FUNCTION_BLOCK FB_PackagingCounter (* Migrated from IEC 61131-3 ST *)
  (* Standard: 61499-2 *)
  (* Version 1.0, 2026-11-06, st2fb *)
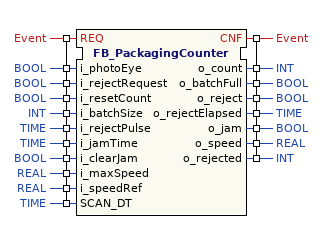
  EVENT_INPUT
    REQ WITH i_photoEye, i_rejectRequest, i_resetCount, i_batchSize, i_rejectPulse, i_jamTime, i_clearJam, i_maxSpeed, i_speedRef, SCAN_DT;
  END_EVENT
  EVENT_OUTPUT
    CNF WITH o_count, o_batchFull, o_reject, o_rejectElapsed, o_jam, o_speed, o_rejected;
  END_EVENT
  VAR_INPUT
    i_photoEye : BOOL;
    i_rejectRequest : BOOL;
    i_resetCount : BOOL;
    i_batchSize : INT;
    i_rejectPulse : TIME;
    i_jamTime : TIME;
    i_clearJam : BOOL;
    i_maxSpeed : REAL;
    i_speedRef : REAL;
    SCAN_DT : TIME;
  END_VAR
  VAR_OUTPUT
    o_count : INT;
    o_batchFull : BOOL;
    o_reject : BOOL;
    o_rejectElapsed : TIME;
    o_jam : BOOL;
    o_speed : REAL;
    o_rejected : INT;
  END_VAR
  VAR
    statEyePrev : BOOL := FALSE;
    statRequestPrev : BOOL := FALSE;
    statRejectPrev : BOOL := FALSE;
    statRejectPreset : TIME := T#0s;
    statJamPreset : TIME := T#0s;
    tempCartonEdge : BOOL := FALSE;
    tempRejectEdge : BOOL := FALSE;
    ST2FB_NOW : TIME := T#0s;
    RP_IN : BOOL := FALSE;
    RP_PT : TIME := T#0s;
    RP_Q : BOOL := FALSE;
    RP_ET : TIME := T#0s;
    RP_STATE : INT := 0;
    RP_PREV_IN : BOOL := FALSE;
    RP_START_TIME : TIME := T#0s;
    JT_IN : BOOL := FALSE;
    JT_PT : TIME := T#0s;
    JT_Q : BOOL := FALSE;
    JT_ET : TIME := T#0s;
    JT_STATE : INT := 0;
    JT_PREV_IN : BOOL := FALSE;
    JT_START_TIME : TIME := T#0s;
  END_VAR
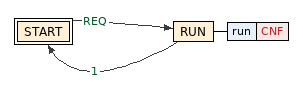
  EC_STATES
    START;
    RUN : run -> CNF;
  END_STATES
  EC_TRANSITIONS
    START TO RUN := REQ;
    RUN TO START := 1;
  END_TRANSITIONS
  ALGORITHM run IN ST:
ST2FB_NOW := ST2FB_NOW + SCAN_DT;

tempCartonEdge := statEyePrev AND NOT i_photoEye;
IF i_resetCount THEN
  o_count := 0;
ELSIF tempCartonEdge AND o_count < i_batchSize THEN
  o_count := o_count + 1;
END_IF;
o_batchFull := o_count >= i_batchSize;

tempRejectEdge := statRequestPrev AND NOT i_rejectRequest;
statRequestPrev := i_rejectRequest;
IF NOT o_reject THEN
  statRejectPreset := i_rejectPulse;
END_IF;
RP_IN := tempRejectEdge AND NOT o_jam;
RP_PT := statRejectPreset;
IF (RP_STATE = 0) AND NOT RP_PREV_IN AND RP_IN THEN
  RP_STATE := 1;
  RP_Q := TRUE;
  RP_START_TIME := ST2FB_NOW;
ELSIF RP_STATE = 1 THEN
  IF RP_START_TIME + RP_PT <= ST2FB_NOW THEN
    RP_STATE := 2;
    RP_Q := FALSE;
    RP_ET := RP_PT;
  ELSE
    RP_ET := ST2FB_NOW - RP_START_TIME;
  END_IF;
END_IF;
IF (RP_STATE = 2) AND NOT RP_IN THEN
  RP_ET := T#0s;
  RP_STATE := 0;
END_IF;
RP_PREV_IN := RP_IN;
o_reject := RP_Q;
o_rejectElapsed := RP_ET;
IF i_resetCount THEN
  o_rejected := 0;
ELSIF o_reject AND NOT statRejectPrev THEN
  o_rejected := o_rejected + 1;
END_IF;
statRejectPrev := o_reject;

IF NOT statEyePrev THEN
  statJamPreset := i_jamTime;
END_IF;
statEyePrev := i_photoEye;
JT_IN := i_photoEye;
JT_PT := statJamPreset;
IF (JT_STATE = 0) AND NOT JT_PREV_IN AND JT_IN THEN
  JT_STATE := 1;
  JT_Q := FALSE;
  JT_START_TIME := ST2FB_NOW;
ELSE
  IF NOT JT_IN THEN
    JT_ET := T#0s;
    JT_Q := FALSE;
    JT_STATE := 0;
  ELSIF JT_STATE = 1 THEN
    IF JT_START_TIME + JT_PT <= ST2FB_NOW THEN
      JT_STATE := 2;
      JT_Q := TRUE;
      JT_ET := JT_PT;
    ELSE
      JT_ET := ST2FB_NOW - JT_START_TIME;
    END_IF;
  END_IF;
END_IF;
JT_PREV_IN := JT_IN;
IF JT_Q THEN
  o_jam := TRUE;
ELSIF i_clearJam THEN
  o_jam := FALSE;
END_IF;
IF o_jam OR o_batchFull THEN
  o_speed := 0.0;
ELSE
  o_speed := MIN(i_speedRef, i_maxSpeed);
END_IF;
  END_ALGORITHM
END_FUNCTION_BLOCK
